Staubli VAL3: setAngOUTList.pgx

public program setAngOUTList(string& x_sList[])
  local num l_i
begin
  resize(x_sList,1,nMaxAnalog)
  for l_i = 0 to nMaxAnalog-1
    x_sList[l_i]=toString("",l_i)+","+aOutItem[l_i].sComment
  endFor
end
